// SIMATIC S7-200 project (STEP 7-Micro/WIN), CPU 224XP CN REL 02.01

SYMBOL_TABLE 用户定义1
编码器A             I0.0
编码器B             I0.1
编码器Z             I0.2
物料口检测传感器         I0.3
光纤传感器            I0.4
接近开关             I0.5
推杆一到位检测          I0.7
推杆二到位检测          I1.0
推杆三到位检测          I1.1
确认按钮             I1.2
启动按钮             I1.3
急停按钮             I1.4
单机全线             I1.5
准备就绪             M0.0
启动               M0.1
金属工件             M1.0
铁芯               M1.1
铁芯金属             M1.2
白芯塑料             M1.3
其他               M1.4
变频器启停控制          Q0.0
推料一电磁阀           Q0.4
推料二电磁阀           Q0.5
推料三电磁阀           Q0.6
黄色指示灯            Q0.7
绿色指示灯            Q1.0
红色指示灯            Q1.1
供料请求_主站          V1000.4
允许分拣             V1000.7
全线停止             V1001.0
套件清零             V1001.2
网络正常             V1010.0
全线模式             V1010.1
停止完成             V1010.2
已生产套件数           VB1011
变频器频率设置          VW1002
END_SYMBOL_TABLE

ORGANIZATION_BLOCK 主程序:OB1
TITLE=程序注释
BEGIN
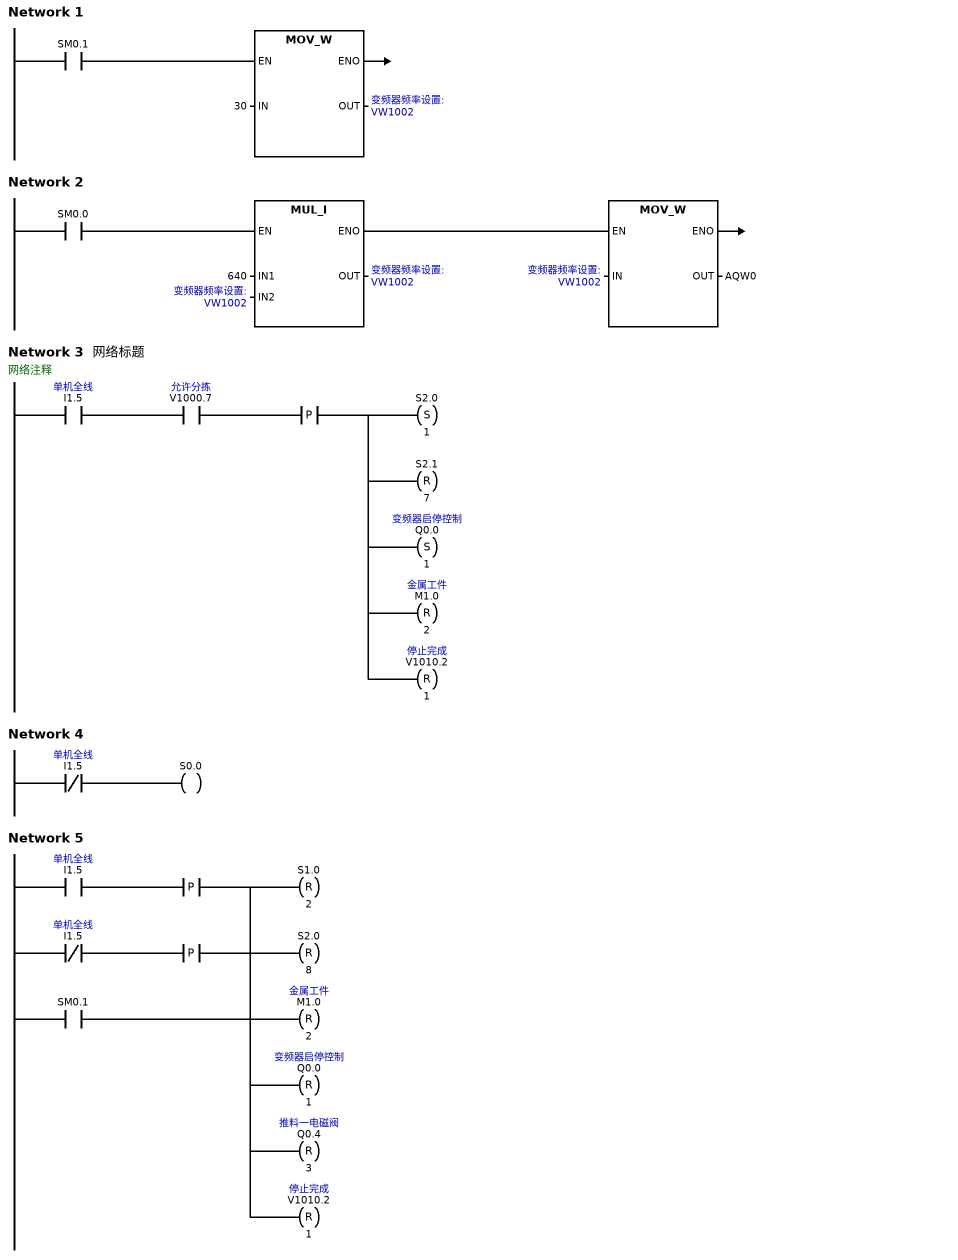
Network 1
LD     SM0.1
MOVW   30, 变频器频率设置:VW1002
Network 2
LD     SM0.0
*I     640, 变频器频率设置:VW1002
AENO
MOVW   变频器频率设置:VW1002, AQW0
Network 3 // 网络标题
// 网络注释
LD     单机全线:I1.5
A      允许分拣:V1000.7
EU
S      S2.0, 1
R      S2.1, 7
S      变频器启停控制:Q0.0, 1
R      金属工件:M1.0, 2
R      停止完成:V1010.2, 1
Network 4
LDN    单机全线:I1.5
=      S0.0
Network 5
LD     单机全线:I1.5
EU
LDN    单机全线:I1.5
EU
OLD
O      SM0.1
R      S1.0, 2
R      S2.0, 8
R      金属工件:M1.0, 2
R      变频器启停控制:Q0.0, 1
R      推料一电磁阀:Q0.4, 3
R      停止完成:V1010.2, 1
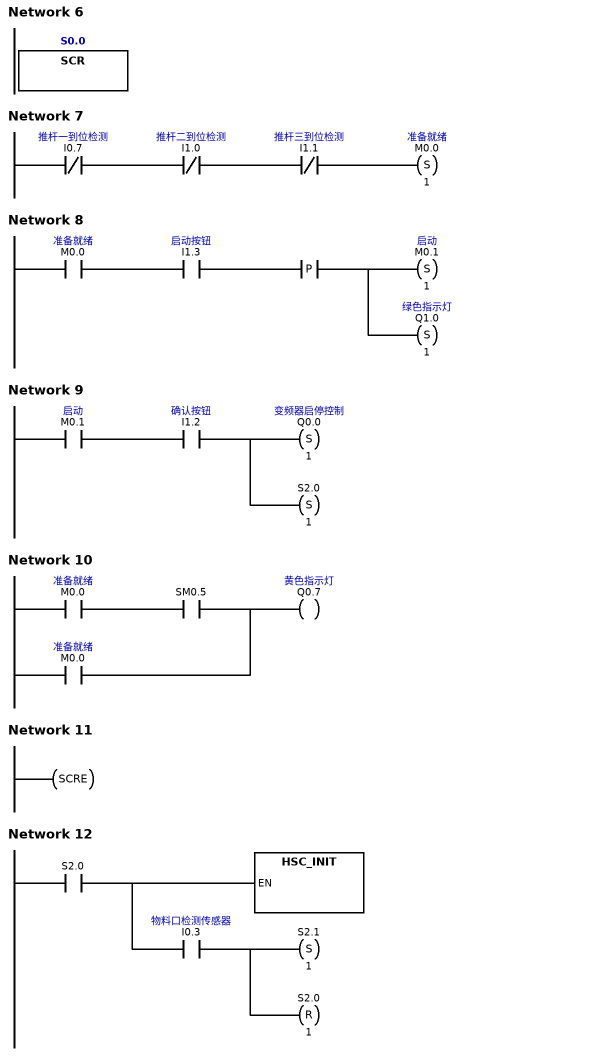
Network 6
LSCR   S0.0
Network 7
LDN    推杆一到位检测:I0.7
AN     推杆二到位检测:I1.0
AN     推杆三到位检测:I1.1
S      准备就绪:M0.0, 1
Network 8
LD     准备就绪:M0.0
A      启动按钮:I1.3
EU
S      启动:M0.1, 1
S      绿色指示灯:Q1.0, 1
Network 9
LD     启动:M0.1
A      确认按钮:I1.2
S      变频器启停控制:Q0.0, 1
S      S2.0, 1
Network 10
LD     准备就绪:M0.0
A      SM0.5
O      准备就绪:M0.0
=      黄色指示灯:Q0.7
Network 11
SCRE
Network 12
LD     S2.0
CALL   HSC_INIT:SBR1
A      物料口检测传感器:I0.3
S      S2.1, 1
R      S2.0, 1
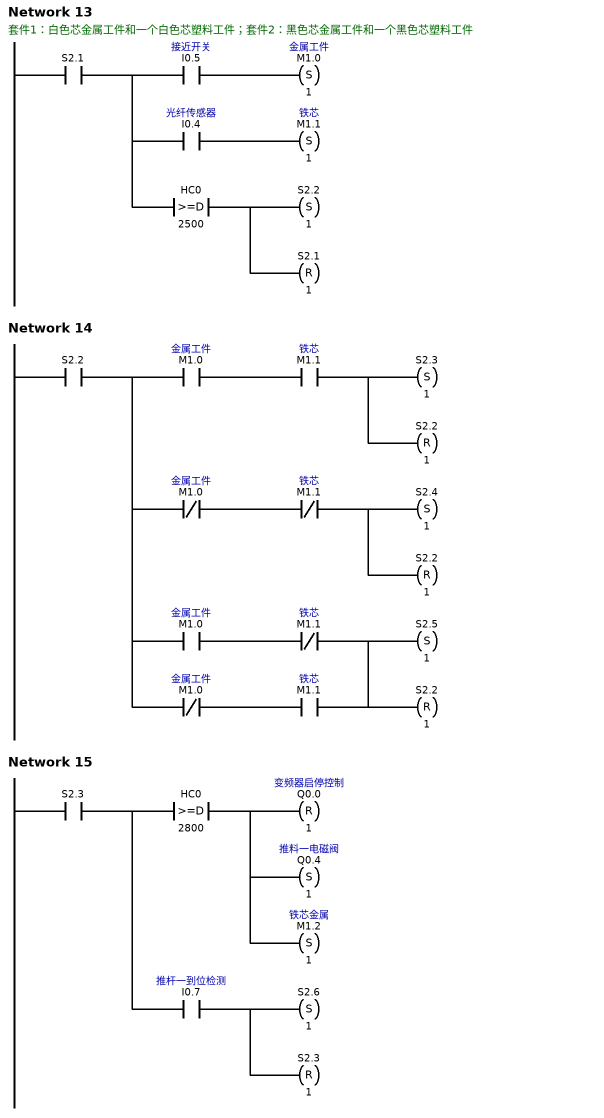
Network 13
// 套件1：白色芯金属工件和一个白色芯塑料工件；套件2：黑色芯金属工件和一个黑色芯塑料工件
LD     S2.1
LPS
A      接近开关:I0.5
S      金属工件:M1.0, 1
LRD
A      光纤传感器:I0.4
S      铁芯:M1.1, 1
LPP
AD>=   HC0, 2500
S      S2.2, 1
R      S2.1, 1
Network 14
LD     S2.2
LPS
A      金属工件:M1.0
A      铁芯:M1.1
S      S2.3, 1
R      S2.2, 1
LRD
AN     金属工件:M1.0
AN     铁芯:M1.1
S      S2.4, 1
R      S2.2, 1
LPP
LD     金属工件:M1.0
AN     铁芯:M1.1
LDN    金属工件:M1.0
A      铁芯:M1.1
OLD
ALD
S      S2.5, 1
R      S2.2, 1
Network 15
LD     S2.3
LPS
AD>=   HC0, 2800
R      变频器启停控制:Q0.0, 1
S      推料一电磁阀:Q0.4, 1
S      铁芯金属:M1.2, 1
LPP
A      推杆一到位检测:I0.7
S      S2.6, 1
R      S2.3, 1
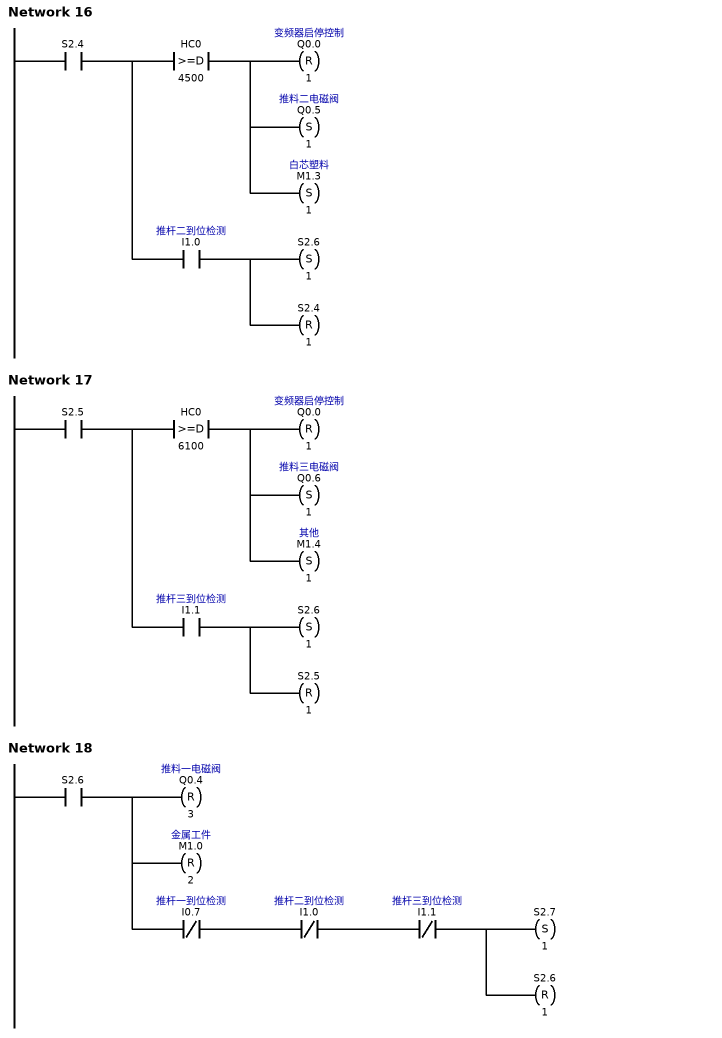
Network 16
LD     S2.4
LPS
AD>=   HC0, 4500
R      变频器启停控制:Q0.0, 1
S      推料二电磁阀:Q0.5, 1
S      白芯塑料:M1.3, 1
LPP
A      推杆二到位检测:I1.0
S      S2.6, 1
R      S2.4, 1
Network 17
LD     S2.5
LPS
AD>=   HC0, 6100
R      变频器启停控制:Q0.0, 1
S      推料三电磁阀:Q0.6, 1
S      其他:M1.4, 1
LPP
A      推杆三到位检测:I1.1
S      S2.6, 1
R      S2.5, 1
Network 18
LD     S2.6
R      推料一电磁阀:Q0.4, 3
R      金属工件:M1.0, 2
AN     推杆一到位检测:I0.7
AN     推杆二到位检测:I1.0
AN     推杆三到位检测:I1.1
S      S2.7, 1
R      S2.6, 1
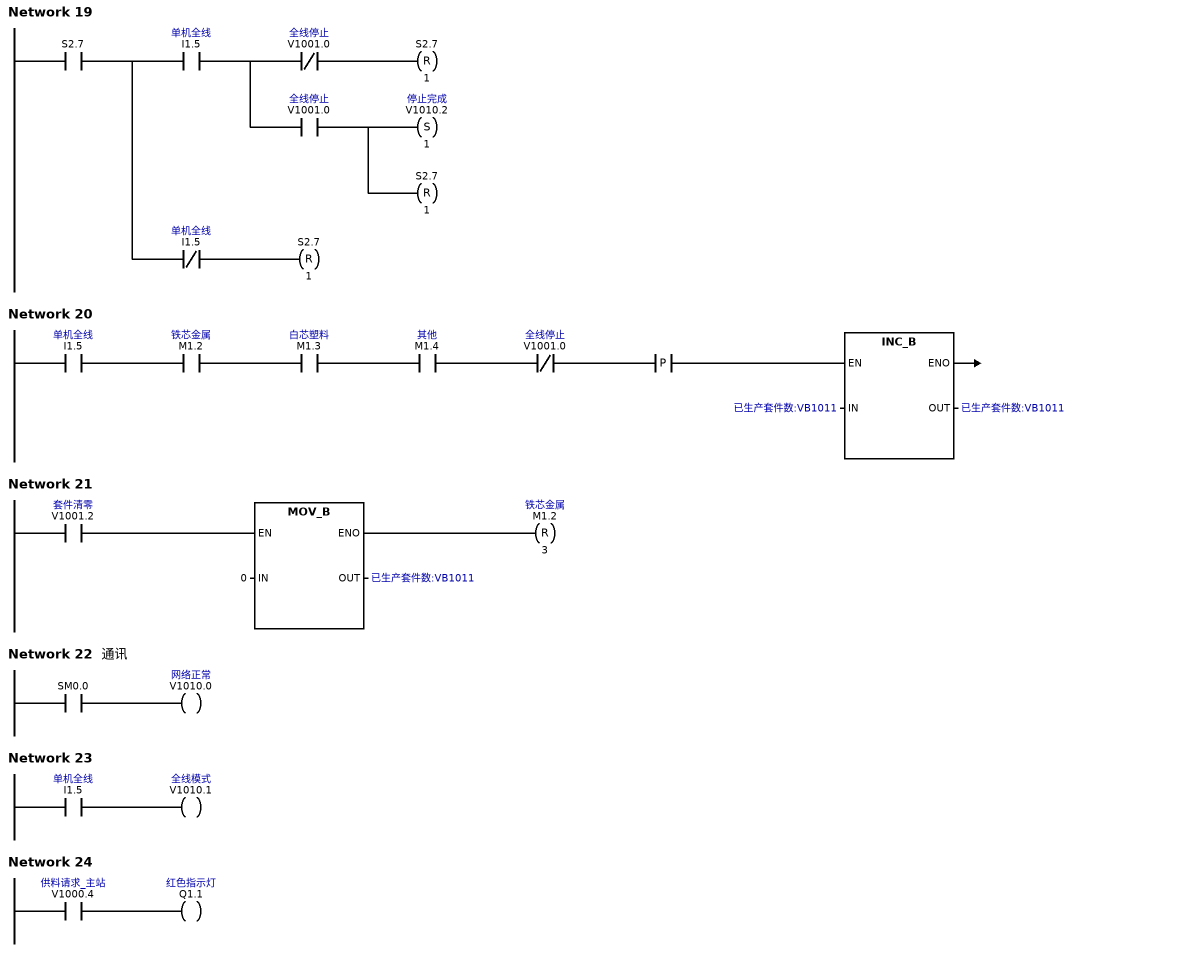
Network 19
LD     S2.7
LPS
A      单机全线:I1.5
LPS
AN     全线停止:V1001.0
R      S2.7, 1
LPP
A      全线停止:V1001.0
S      停止完成:V1010.2, 1
R      S2.7, 1
LPP
AN     单机全线:I1.5
R      S2.7, 1
Network 20
LD     单机全线:I1.5
A      铁芯金属:M1.2
A      白芯塑料:M1.3
A      其他:M1.4
AN     全线停止:V1001.0
EU
INCB   已生产套件数:VB1011
Network 21
LD     套件清零:V1001.2
MOVB   0, 已生产套件数:VB1011
AENO
R      铁芯金属:M1.2, 3
Network 22 // 通讯
LD     SM0.0
=      网络正常:V1010.0
Network 23
LD     单机全线:I1.5
=      全线模式:V1010.1
Network 24
LD     供料请求_主站:V1000.4
=      红色指示灯:Q1.1
END_ORGANIZATION_BLOCK

SUBROUTINE_BLOCK HSC_INIT:SBR1
TITLE=
BEGIN
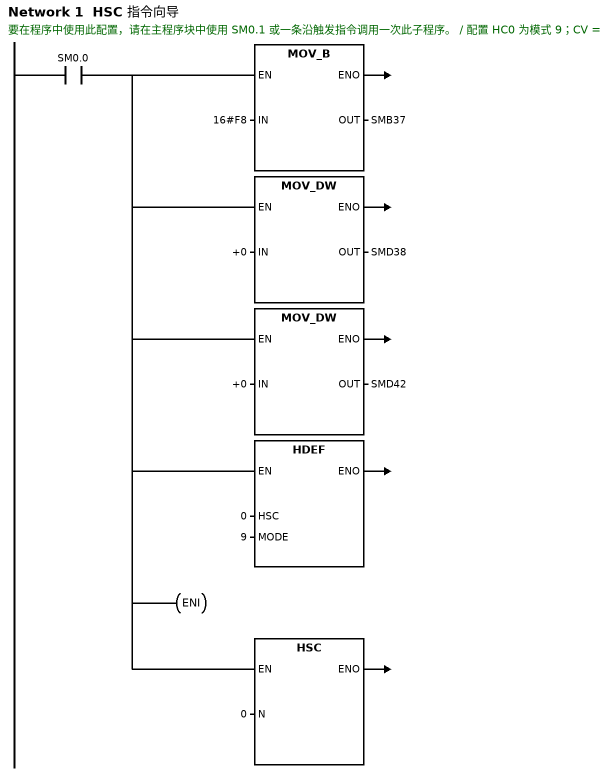
Network 1 // HSC 指令向导
// 要在程序中使用此配置，请在主程序块中使用 SM0.1 或一条沿触发指令调用一次此子程序。
// 配置 HC0 为模式 9；CV = 0； PV = 0；增计数；
// 开放中断和启动计数器。
// 
//设置控制位：增计数；4X 速率；已使能；
//装载 CV
//装载 PV
LD     SM0.0
MOVB   16#F8, SMB37
MOVD   +0, SMD38
MOVD   +0, SMD42
HDEF   0, 9
ENI
HSC    0
END_SUBROUTINE_BLOCK
